(* IEC 61131-3 sources: kns-pump-station/tests/POUs/Station/FB_LevelControlStepped_Test, 13 files *)

(* ---- AssistOnAndOffWithHysteresis.method.decl.st ---- *)
// 04 §6, PMI-03: подпорный — пуск при 2,40 м, между 1,40 и 2,40 м число держится, останов подпорного при 1,40 м;
// ведущий работает выше 1,00 м
METHOD PRIVATE AssistOnAndOffWithHysteresis
VAR
    fbDut  : FB_LevelControlStepped;    // ФБ под тестом
    fbTime : PL.FB_FakeTime;            // подменное время, старт 1 ч
    stCfg  : ST_StationCfg;             // уставки по умолчанию (04 §18.2)
END_VAR

(* ---- BoundaryLevelsInclusive.method.decl.st ---- *)
// 04 §6: границы включительно — пуск подпорного ровно при 2,40 м, останов подпорного ровно при 1,40 м; 1,59 м —
// без пуска
METHOD PRIVATE BoundaryLevelsInclusive
VAR
    fbDut  : FB_LevelControlStepped;    // ФБ под тестом
    fbTime : PL.FB_FakeTime;            // подменное время, старт 1 ч
    stCfg  : ST_StationCfg;             // уставки по умолчанию (04 §18.2)
    fbDut2 : FB_LevelControlStepped;   // второй экземпляр: уровень чуть ниже пуска
END_VAR

(* ---- DisabledOutputsZeroInitRestores.method.decl.st ---- *)
// DESIGN 6.3: xEnable = FALSE — выход 0, автомат продолжает работу; следующий xInit задаёт состояние по работающим
METHOD PRIVATE DisabledOutputsZeroInitRestores
VAR
    fbDut  : FB_LevelControlStepped;    // ФБ под тестом
    fbTime : PL.FB_FakeTime;            // подменное время, старт 1 ч
    stCfg  : ST_StationCfg;             // уставки по умолчанию (04 §18.2)
END_VAR

(* ---- DutyMaxOneLimitsToOne.method.decl.st ---- *)
// 04 §18.2 № 13: uiDutyMax = 1 — не больше одного насоса и при инициализации, и выше уровня пуска подпорного
METHOD PRIVATE DutyMaxOneLimitsToOne
VAR
    fbDut  : FB_LevelControlStepped;    // ФБ под тестом
    fbTime : PL.FB_FakeTime;            // подменное время, старт 1 ч
    stCfg  : ST_StationCfg;             // уставки по умолчанию (04 §18.2)
END_VAR

(* ---- InitFromRunningPumpsNoStop.method.decl.st ---- *)
// 04 §3.2, PMI-07: вход без рывка — число насосов по работающим, при уровне между остановом и пуском насос не
// останавливается
METHOD PRIVATE InitFromRunningPumpsNoStop
VAR
    fbDut  : FB_LevelControlStepped;    // ФБ под тестом
    fbTime : PL.FB_FakeTime;            // подменное время, старт 1 ч
    stCfg  : ST_StationCfg;             // уставки по умолчанию (04 §18.2)
END_VAR

(* ---- InvalidLevelHoldsState.method.decl.st ---- *)
// 04 §6: недостоверный уровень (и NaN при xLevelValid) — число насосов держится, выдержки не идут
METHOD PRIVATE InvalidLevelHoldsState
VAR
    fbDut  : FB_LevelControlStepped;    // ФБ под тестом
    fbTime : PL.FB_FakeTime;            // подменное время, старт 1 ч
    stCfg  : ST_StationCfg;             // уставки по умолчанию (04 §18.2)
    rNan   : REAL;                     // NaN
    uBits  : PL.U_RealBits;             // сборка NaN по битам
END_VAR

(* ---- NoStartIfLevelDropsDuringConfirm.method.decl.st ---- *)
// 04 §6: волна — уровень опустился ниже пуска до конца выдержки: пуска нет, выдержка начинается заново
METHOD PRIVATE NoStartIfLevelDropsDuringConfirm
VAR
    fbDut  : FB_LevelControlStepped;    // ФБ под тестом
    fbTime : PL.FB_FakeTime;            // подменное время, старт 1 ч
    stCfg  : ST_StationCfg;             // уставки по умолчанию (04 §18.2)
END_VAR

(* ---- Run.method.decl.st ---- *)
// Помощник: uiSteps шагов по 100 мс с одним уровнем; в каждом шаге — сначала время, потом вызов
METHOD PRIVATE Run
VAR_IN_OUT
    fbDut  : FB_LevelControlStepped;    // ФБ под тестом
    fbTime : PL.FB_FakeTime;            // подменное время
    stCfg  : ST_StationCfg;             // уставки
END_VAR
VAR_INPUT
    rLevel_m : REAL;                    // уровень
    xValid   : BOOL;                    // уровень достоверен
    uiSteps  : UINT;                    // шагов по 100 мс
END_VAR
VAR
    uiStep : UINT;                      // номер шага
END_VAR

(* ---- Run.method.impl.st ---- *)
FOR uiStep := 1 TO uiSteps DO
    fbTime.Advance(tStep := T#100MS);
    fbDut(xEnable := TRUE, rLevel_m := rLevel_m, xLevelValid := xValid, xInit := FALSE, itfTime := fbTime,
          stCfg := stCfg);
END_FOR

(* ---- StartsLeadAtStartLevelAfterConfirm.method.decl.st ---- *)
// 04 §6, PMI-02: уровень 1,60 м (граница пуска ведущего) — пуск ровно через tLvlConfirm = 5 с, не на шаге раньше;
// частота — rStepSpeed_pct
METHOD PRIVATE StartsLeadAtStartLevelAfterConfirm
VAR
    fbDut  : FB_LevelControlStepped;    // ФБ под тестом
    fbTime : PL.FB_FakeTime;            // подменное время, старт 1 ч
    stCfg  : ST_StationCfg;             // уставки по умолчанию (04 §18.2)
END_VAR

(* ---- StopsAllAtStopLevel.method.decl.st ---- *)
// 04 §6, PMI-02: один насос, уровень 1,00 м (граница останова) — останов ровно через 5 с
METHOD PRIVATE StopsAllAtStopLevel
VAR
    fbDut  : FB_LevelControlStepped;    // ФБ под тестом
    fbTime : PL.FB_FakeTime;            // подменное время, старт 1 ч
    stCfg  : ST_StationCfg;             // уставки по умолчанию (04 §18.2)
END_VAR

(* ---- TimeBackwardsRestartsConfirm.method.decl.st ---- *)
// Время назад (сбой источника) — выдержка подтверждения начинается заново, ложного пуска нет
METHOD PRIVATE TimeBackwardsRestartsConfirm
VAR
    fbDut  : FB_LevelControlStepped;    // ФБ под тестом
    fbTime : PL.FB_FakeTime;            // подменное время, старт 1 ч
    stCfg  : ST_StationCfg;             // уставки по умолчанию (04 §18.2)
END_VAR

(* ---- TwoToZeroAtStopLevel.method.decl.st ---- *)
// 04 §6: два насоса, уровень сразу ниже останова — оба останавливаются одним переходом через 5 с
METHOD PRIVATE TwoToZeroAtStopLevel
VAR
    fbDut  : FB_LevelControlStepped;    // ФБ под тестом
    fbTime : PL.FB_FakeTime;            // подменное время, старт 1 ч
    stCfg  : ST_StationCfg;             // уставки по умолчанию (04 §18.2)
END_VAR
